DATA_BLOCK "FRK_SetStore"
{ S7_Optimized_Access := 'TRUE' }
VERSION : 0.1
NON_RETAIN
VAR RETAIN
    SchemaVersion {ExternalAccessible := 'False'; ExternalVisible := 'False'; ExternalWritable := 'False'} : UInt;
    Sets {ExternalAccessible := 'False'; ExternalVisible := 'False'; ExternalWritable := 'False'} : Array[1..2, 1..4] of "FRK_SetPayload";
END_VAR
BEGIN
END_DATA_BLOCK
